// TIA Portal V20 export
// export: Created 2026-10-12T05:42:35.6266844Z, ExportSetting WithDefaults, DisplayName Totally Integrated Automation Portal, DisplayVersion V20, DisplayName TIA Portal Openness, DisplayVersion V20, DisplayName TIA Portal Teamcenter Gateway, DisplayVersion V20, DisplayName TIA Portal Version Control Interface, DisplayVersion V20, DisplayName SINAMICS Startdrive Advanced, DisplayVersion V20 SP1 Update 2, DisplayName SINAMICS Startdrive G110M, G120, G120C, G120D, G120P, G115D, DisplayVersion V20 SP1 Update 2, DisplayName SINAMICS Startdrive G130, G150, S120, S150, SINAMICS MV, G220, S200, S210, DisplayVersion V20 SP1 Update 2, DisplayName STEP 7 Professional, DisplayVersion V20, DisplayName STEP 7 Safety, DisplayVersion V20, DisplayName WinCC Basic/Comfort/Advanced, DisplayVersion V20, DisplayName WinCC Professional, DisplayVersion V20, DisplayName WinCC Unified, DisplayVersion V20
FUNCTION_BLOCK "FB_LD_PressDemoRelease"   // FB9, LAD
{ S7_Optimized_Access := 'TRUE' }
VERSION : 0.1
// stored: AutoNumber true, IsIECCheckEnabled false, IsRetainMemResEnabled false, MemoryReserve 100, SetENOAutomatically false, UDAEnableTagReadback false
   VAR_INPUT
      AirPressureOk { ExternalWritable := 'False'} : Bool;
      DoorClosed { ExternalWritable := 'False'} : Bool;
      DoorHealthy { ExternalWritable := 'False'} : Bool;
      RamHealthy { ExternalWritable := 'False'} : Bool;
      SlideHealthy { ExternalWritable := 'False'} : Bool;
      SlideInside { ExternalWritable := 'False'} : Bool;
      TwoHandHeld { ExternalWritable := 'False'} : Bool;
   END_VAR
   VAR
      Conditions { ExternalWritable := 'False'} : "ST_PressDemoReleaseConditions";
      ModeStart { ExternalWritable := 'False'} : "FRK_PermCtx";
      RamExtend { ExternalWritable := 'False'} : "FRK_PermCtx";
   END_VAR
BEGIN

REGION Network 1
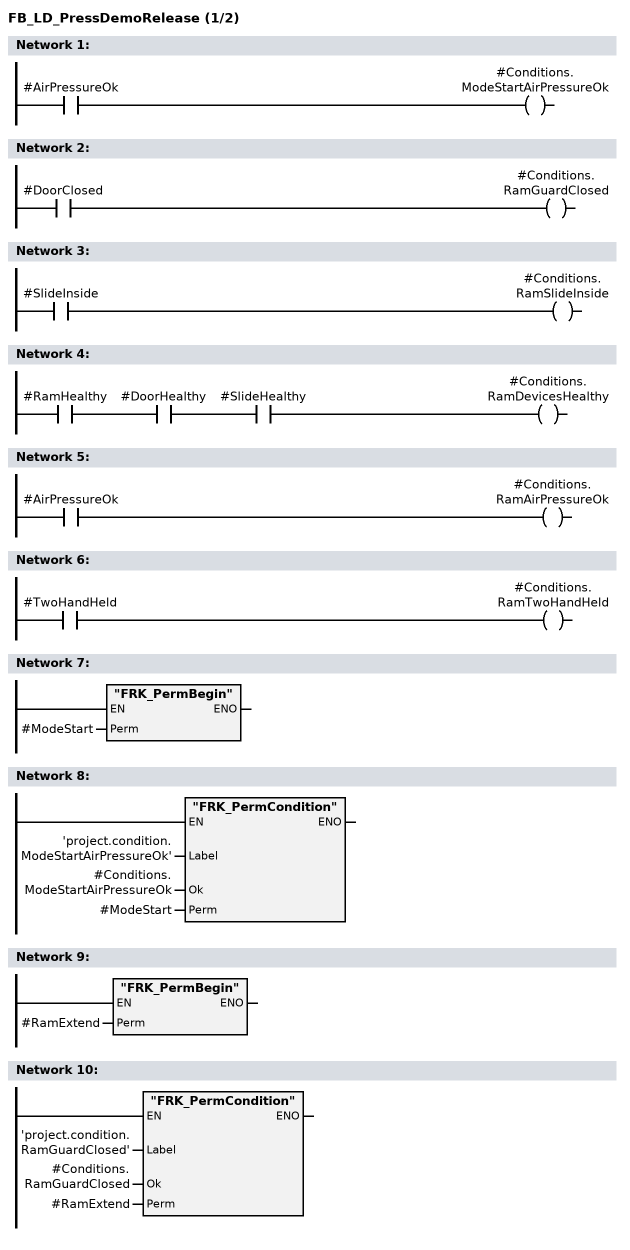
   RUNG wire#powerrail
      Contact( #AirPressureOk )
      Coil( #Conditions.ModeStartAirPressureOk )
   END_RUNG
   // the same network as SCL:
   #Conditions.ModeStartAirPressureOk := #AirPressureOk;
END_REGION

REGION Network 2
   RUNG wire#powerrail
      Contact( #DoorClosed )
      Coil( #Conditions.RamGuardClosed )
   END_RUNG
   // the same network as SCL:
   #Conditions.RamGuardClosed := #DoorClosed;
END_REGION

REGION Network 3
   RUNG wire#powerrail
      Contact( #SlideInside )
      Coil( #Conditions.RamSlideInside )
   END_RUNG
   // the same network as SCL:
   #Conditions.RamSlideInside := #SlideInside;
END_REGION

REGION Network 4
   RUNG wire#powerrail
      Contact( #RamHealthy )
      Contact( #DoorHealthy )
      Contact( #SlideHealthy )
      Coil( #Conditions.RamDevicesHealthy )
   END_RUNG
   // the same network as SCL:
   #Conditions.RamDevicesHealthy := #RamHealthy AND #DoorHealthy AND #SlideHealthy;
END_REGION

REGION Network 5
   RUNG wire#powerrail
      Contact( #AirPressureOk )
      Coil( #Conditions.RamAirPressureOk )
   END_RUNG
   // the same network as SCL:
   #Conditions.RamAirPressureOk := #AirPressureOk;
END_REGION

REGION Network 6
   RUNG wire#powerrail
      Contact( #TwoHandHeld )
      Coil( #Conditions.RamTwoHandHeld )
   END_RUNG
   // the same network as SCL:
   #Conditions.RamTwoHandHeld := #TwoHandHeld;
END_REGION

REGION Network 7
   RUNG wire#powerrail
      "FRK_PermBegin"(Perm := #ModeStart)
   END_RUNG
   // the same network as SCL:
   "FRK_PermBegin"(Perm := #ModeStart);
END_REGION

REGION Network 8
   RUNG wire#powerrail
      "FRK_PermCondition"(Label := 'project.condition.ModeStartAirPressureOk', Ok := #Conditions.ModeStartAirPressureOk, Perm := #ModeStart)
   END_RUNG
   // the same network as SCL:
   "FRK_PermCondition"(Label := 'project.condition.ModeStartAirPressureOk',
                       Ok := #Conditions.ModeStartAirPressureOk,
                       Perm := #ModeStart);
END_REGION

REGION Network 9
   RUNG wire#powerrail
      "FRK_PermBegin"(Perm := #RamExtend)
   END_RUNG
   // the same network as SCL:
   "FRK_PermBegin"(Perm := #RamExtend);
END_REGION

REGION Network 10
   RUNG wire#powerrail
      "FRK_PermCondition"(Label := 'project.condition.RamGuardClosed', Ok := #Conditions.RamGuardClosed, Perm := #RamExtend)
   END_RUNG
   // the same network as SCL:
   "FRK_PermCondition"(Label := 'project.condition.RamGuardClosed',
                       Ok := #Conditions.RamGuardClosed,
                       Perm := #RamExtend);
END_REGION

REGION Network 11
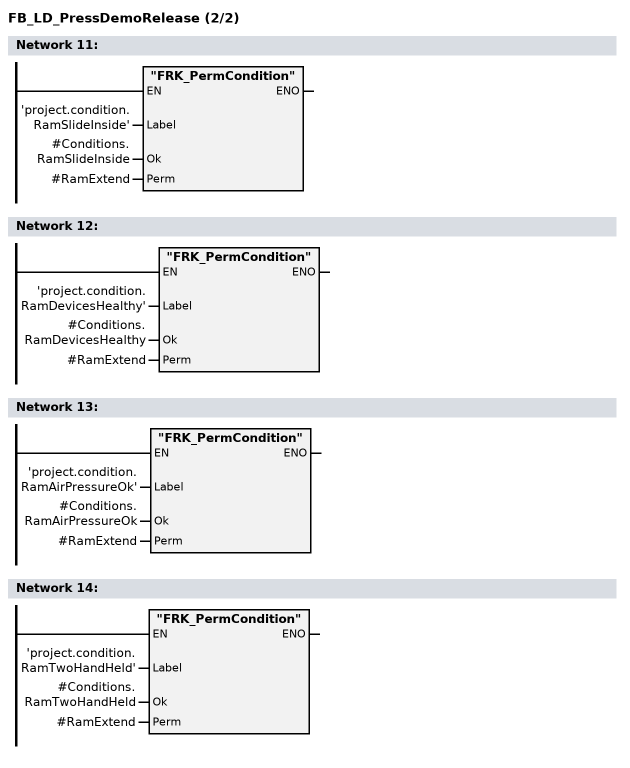
   RUNG wire#powerrail
      "FRK_PermCondition"(Label := 'project.condition.RamSlideInside', Ok := #Conditions.RamSlideInside, Perm := #RamExtend)
   END_RUNG
   // the same network as SCL:
   "FRK_PermCondition"(Label := 'project.condition.RamSlideInside',
                       Ok := #Conditions.RamSlideInside,
                       Perm := #RamExtend);
END_REGION

REGION Network 12
   RUNG wire#powerrail
      "FRK_PermCondition"(Label := 'project.condition.RamDevicesHealthy', Ok := #Conditions.RamDevicesHealthy, Perm := #RamExtend)
   END_RUNG
   // the same network as SCL:
   "FRK_PermCondition"(Label := 'project.condition.RamDevicesHealthy',
                       Ok := #Conditions.RamDevicesHealthy,
                       Perm := #RamExtend);
END_REGION

REGION Network 13
   RUNG wire#powerrail
      "FRK_PermCondition"(Label := 'project.condition.RamAirPressureOk', Ok := #Conditions.RamAirPressureOk, Perm := #RamExtend)
   END_RUNG
   // the same network as SCL:
   "FRK_PermCondition"(Label := 'project.condition.RamAirPressureOk',
                       Ok := #Conditions.RamAirPressureOk,
                       Perm := #RamExtend);
END_REGION

REGION Network 14
   RUNG wire#powerrail
      "FRK_PermCondition"(Label := 'project.condition.RamTwoHandHeld', Ok := #Conditions.RamTwoHandHeld, Perm := #RamExtend)
   END_RUNG
   // the same network as SCL:
   "FRK_PermCondition"(Label := 'project.condition.RamTwoHandHeld',
                       Ok := #Conditions.RamTwoHandHeld,
                       Perm := #RamExtend);
END_REGION
END_FUNCTION_BLOCK
